(* PLC project CIP_Plant.project, CODESYS CODESYS V3.5 SP22 Patch 4 *)
(* stored: creationDateTime 2026-10-20T09:44:48.4195395, modificationDateTime 2026-10-20T09:30:51.2284783 *)

PROGRAM PLC_PRG
VAR
	Start_Btn : BOOL;
	Valve_Out : BOOL;
Delay : TON;
END_VAR

             Delay(IN := Start_Btn, PT := T#5S);
Valve_Out := Delay.Q;
 
          
END_PROGRAM
